(* IEC 61131-3 sources: volt/packages/volt-lsp-iec/test-corpus/bakon-nano/Device/Plc Logic/Application/Library Manager/Collections, 40 files *)

(* ---- PAIR_DINTDINT.dut ---- *)
TYPE PAIR_DINTDINT :
STRUCT
	DIKEY : DINT;
	DIVALUE : DINT;
END_STRUCT
END_TYPE

(* ---- PAIR_PSTRINGDINT.dut ---- *)
TYPE PAIR_PSTRINGDINT :
STRUCT
	PSTR : POINTER TO STRING;
	DI : DINT;
END_STRUCT
END_TYPE

(* ---- PAIR_PSTRINGXWORD.dut ---- *)
TYPE PAIR_PSTRINGXWORD :
STRUCT
	PSTR : POINTER TO STRING;
	XW : __XWORD;
END_STRUCT
END_TYPE

(* ---- PAIR_STRINGDINT.dut ---- *)
TYPE PAIR_STRINGDINT :
STRUCT
	STR : STRING;
	DI : DINT;
END_STRUCT
END_TYPE

(* ---- PAIR_STRINGSTRING.dut ---- *)
TYPE PAIR_STRINGSTRING :
STRUCT
	STRKEY : STRING;
	STRVALUE : STRING;
END_STRUCT
END_TYPE

(* ---- STATICMEMBUFFER.dut ---- *)
TYPE STATICMEMBUFFER :
STRUCT
	PDATA : POINTER TO BYTE;
	UDIDATASIZE : UDINT;
	XEXTENDDYNAMICALLY : BOOL;
END_STRUCT
END_TYPE

(* ---- GLOBALS.gvl ---- *)
VAR_GLOBAL
	COMPONENT_NAME : STRING := 'Collections';
	VECTOR_STRING_LEN : INT := 80;
	ERR_MB_ALREADY_ALLOCATED : UDINT := 16#2100;
	ERR_OK : UDINT := 0;
	ERR_PARAMETER : UDINT := 2;
	ERR_NOTINITIALIZED : UDINT := 3;
	ERR_NOBUFFER : UDINT := 6;
	ERR_NOTIMPLEMENTED : UDINT := 12;
	ERR_NO_OBJECT : UDINT := 16#16;
END_VAR

(* ---- GVL_DEBUGONLYCOLLECTIONS.gvl ---- *)
VAR_GLOBAL
	G_ST : STRING(255);
	G_PST : POINTER TO STRING(255);
END_VAR

(* ---- PSTRCAT.pou ---- *)
FUNCTION PSTRCAT : DINT
VAR_INPUT
	PSTDEST : POINTER TO STRING;
	PSTSRC : POINTER TO STRING;
	DIDESTSIZE : DINT;
END_VAR
END_FUNCTION

(* ---- PSTRCMP.pou ---- *)
FUNCTION PSTRCMP : INT
VAR_INPUT
	PSTR1 : POINTER TO STRING;
	PSTR2 : POINTER TO STRING;
END_VAR
END_FUNCTION

(* ---- PSTRICMP.pou ---- *)
FUNCTION PSTRICMP : INT
VAR_INPUT
	PSTR1 : POINTER TO STRING;
	PSTR2 : POINTER TO STRING;
END_VAR
END_FUNCTION

(* ---- PSTRIFIND.pou ---- *)
FUNCTION PSTRIFIND : INT
VAR_INPUT
	PST1 : POINTER TO STRING(255);
	PST2 : POINTER TO STRING(255);
END_VAR
END_FUNCTION

(* ---- PSTRLEN.pou ---- *)
FUNCTION PSTRLEN : DINT
VAR_INPUT
	PSTRING : POINTER TO STRING;
END_VAR
END_FUNCTION

(* ---- PSTRLENUNTIL.pou ---- *)
FUNCTION PSTRLENUNTIL : DINT
VAR_INPUT
	PST : POINTER TO STRING;
	STTOKENDELIMITERS : STRING;
END_VAR
END_FUNCTION

(* ---- PSTRTOUPPER.pou ---- *)
FUNCTION PSTRTOUPPER : STRING(255)
VAR_INPUT
	PSTVALUE : POINTER TO STRING(255);
END_VAR
END_FUNCTION

(* ---- ABSTRTREENODE.pou ---- *)
FUNCTION_BLOCK ABSTRTREENODE
VAR
	_FATHER : IBaseTreeNode;
	_ICOUNT : DINT;
	_IBASETREENODE : IBaseTreeNode;
	ABSTRNODETYPE : INT;
	CHILDCOUNT : DINT;
	PROCHILDREN : POINTER TO ARRAY [0..100] OF IBaseTreeNode;
	SORTED : BOOL;
END_VAR
END_FUNCTION_BLOCK

METHOD GETCHILD : IBaseTreeNode
VAR_INPUT
	DIINDEX : DINT;
END_VAR
END_METHOD

METHOD GETFATHER : IBaseTreeNode
END_METHOD

METHOD ABSTRCOMPARETO : INT
VAR_INPUT
	PSEARCHDATA : POINTER TO BYTE;
END_VAR
END_METHOD

METHOD PROFINDCHILDINDEX : DINT
VAR_INPUT
	PSEARCHDATA : POINTER TO BYTE;
END_VAR
END_METHOD

METHOD PROGETNODE : IBaseTreeNode
VAR_INPUT
	DIINDEX : DINT;
END_VAR
END_METHOD

METHOD PRVFINDBINARY : DINT
VAR_INPUT
	PSEARCHDATA : POINTER TO BYTE;
END_VAR
END_METHOD

METHOD PRVFINDLINEAR : DINT
VAR_INPUT
	PSEARCHDATA : POINTER TO BYTE;
END_VAR
END_METHOD

METHOD ADDREF : DINT
END_METHOD

METHOD FB_EXIT : BOOL
VAR_INPUT
	BINCOPYCODE : BOOL;
END_VAR
END_METHOD

METHOD FB_INIT : BOOL
VAR_INPUT
	BINITRETAINS : BOOL;
	BINCOPYCODE : BOOL;
END_VAR
END_METHOD

METHOD FB_REINIT : BOOL
END_METHOD

METHOD QUERYINTERFACE : POINTER TO POINTER TO BYTE
VAR_INPUT
	IID : DWORD;
	PRESULT : POINTER TO UDINT;
END_VAR
END_METHOD

METHOD RELEASE : DINT
END_METHOD

(* ---- BASEMAP.pou ---- *)
FUNCTION_BLOCK BASEMAP EXTENDS BaseVector
VAR
	_IUPDATECOUNT : INT;
	_BOPTIMIZEDSORTFORINSERTIONONLYATEND : BOOL;
	PROUSEOPTIMIZEDSORTFORINSERTIONATTHEEND : BOOL;
END_VAR
END_FUNCTION_BLOCK

METHOD BEGINUPDATE : UDINT
END_METHOD

METHOD ENDUPDATE : UDINT
END_METHOD

METHOD ABSTRCOMPARE : INT
VAR_INPUT
	PKEY1 : POINTER TO BYTE;
	PKEY2 : POINTER TO BYTE;
END_VAR
END_METHOD

METHOD ABSTRKEYPTRFROMINDEX : POINTER TO BYTE
VAR_INPUT
	UDIINDEX : UDINT;
END_VAR
END_METHOD

METHOD ABSTRSWAP : UDINT
VAR_INPUT
	INDEX1 : UDINT;
	INDEX2 : UDINT;
END_VAR
END_METHOD

METHOD PROADDMAPITEM : UDINT
VAR_INPUT
	PITEM : POINTER TO BYTE;
END_VAR
END_METHOD

METHOD PROFINDPAIRINDEX : DINT
VAR_INPUT
	PKEY : POINTER TO BYTE;
END_VAR
END_METHOD

METHOD PRVAFTERUPDATE : UDINT
VAR_INPUT
	BONLYSINGLEINSERT : BOOL;
END_VAR
END_METHOD

METHOD PRVBUBBLESORT : UDINT
END_METHOD

METHOD PRVCOMPAREBYINDEXANDVALUE : INT
VAR_INPUT
	UDI1 : UDINT;
	PKEYVAL : POINTER TO BYTE;
END_VAR
END_METHOD

METHOD PRVCOMPAREBYINDICES : INT
VAR_INPUT
	UDI1 : UDINT;
	UDI2 : UDINT;
END_VAR
END_METHOD

METHOD PRVINSERTIONSORTFORLAST : UDINT
END_METHOD

METHOD PRVSORT : UDINT
VAR_INPUT
	BONLYSINGLEINSERT : BOOL;
END_VAR
END_METHOD

(* ---- BASEVECTOR.pou ---- *)
FUNCTION_BLOCK BASEVECTOR
VAR
	_MEMORY : MemBuffer;
	_PDATA : POINTER TO ARRAY [0..100] OF DWORD;
	_DICURRENTALLOCSIZE : DINT;
	_DICURRENTINSERTPOSITION : DINT;
	CAPACITY : DINT;
	COUNT : DINT;
	PRODATAPTR : POINTER TO BYTE;
END_VAR
END_FUNCTION_BLOCK

METHOD CLEAR : UDINT
END_METHOD

METHOD INITMEMORY : UDINT
VAR_INPUT
	BUFFER : StaticMemBuffer;
END_VAR
END_METHOD

METHOD REMOVELAST : UDINT
END_METHOD

METHOD RESERVESPACE : UDINT
VAR_INPUT
	IITEMCOUNT : UDINT;
END_VAR
END_METHOD

METHOD ABSTRASSIGN : UDINT
VAR_INPUT
	PBT : POINTER TO BYTE;
	UDIINDEX : UDINT;
END_VAR
END_METHOD

METHOD ABSTRDATAPTRCHANGED : UDINT
END_METHOD

METHOD ABSTRGETELEMENTPTR : UDINT
VAR_INPUT
	UDIINDEX : UDINT;
END_VAR
VAR_OUTPUT
	PENTRY : POINTER TO BYTE;
END_VAR
END_METHOD

METHOD ABSTRSIZEOFELEMENT : UDINT
END_METHOD

METHOD PROADDITEM : UDINT
VAR_INPUT
	PBT : POINTER TO BYTE;
END_VAR
END_METHOD

METHOD PROAFTERALLOC
VAR_INPUT
	DIPREVALLOCSIZE : DINT;
	DICURRALLOCSIZE : DINT;
END_VAR
END_METHOD

METHOD PROREMOVE : UDINT
VAR_INPUT
	UDIINDEX : UDINT;
END_VAR
END_METHOD

METHOD PRVALLOC : UDINT
VAR_INPUT
	UDIITEMCOUNT : UDINT;
END_VAR
END_METHOD

(* ---- BRANCHNAMEDTREENODE.pou ---- *)
FUNCTION_BLOCK BRANCHNAMEDTREENODE EXTENDS NamedTreeNode
VAR
	_PCHILDREN : POINTER TO ARRAY [0..100] OF IBaseTreeNode;
	_ICHILDCOUNT : DINT;
	CHILDCOUNT : DINT;
	PROCHILDREN : POINTER TO ARRAY [0..100] OF IBaseTreeNode;
END_VAR
END_FUNCTION_BLOCK

(* ---- CASESENSITIVENAMEDTREENODE.pou ---- *)
FUNCTION_BLOCK CASESENSITIVENAMEDTREENODE EXTENDS NamedTreeNode
VAR
	CASESENSITIVECOMPARISON : BOOL;
END_VAR
END_FUNCTION_BLOCK

(* ---- DINTTODINTMAP.pou ---- *)
FUNCTION_BLOCK DINTTODINTMAP EXTENDS BaseMap
VAR
	_PITEMS : POINTER TO ARRAY [0..100] OF Pair_DintDint;
END_VAR
END_FUNCTION_BLOCK

METHOD ADDDINTPAIR : UDINT
VAR_INPUT
	DIKEY : DINT;
	DIVALUE : DINT;
END_VAR
END_METHOD

METHOD GETVALUE : DINT
VAR_INPUT
	DIKEY : DINT;
END_VAR
VAR_OUTPUT
	UDIRESULT : UDINT;
END_VAR
END_METHOD

METHOD ABSTRASSIGN : UDINT
VAR_INPUT
	PBT : POINTER TO BYTE;
	UDIINDEX : UDINT;
END_VAR
END_METHOD

METHOD ABSTRCOMPARE : INT
VAR_INPUT
	PKEY1 : POINTER TO BYTE;
	PKEY2 : POINTER TO BYTE;
END_VAR
END_METHOD

METHOD ABSTRDATAPTRCHANGED : UDINT
END_METHOD

METHOD ABSTRKEYPTRFROMINDEX : POINTER TO BYTE
VAR_INPUT
	UDIINDEX : UDINT;
END_VAR
END_METHOD

METHOD ABSTRSIZEOFELEMENT : UDINT
END_METHOD

METHOD ABSTRSWAP : UDINT
VAR_INPUT
	INDEX1 : UDINT;
	INDEX2 : UDINT;
END_VAR
END_METHOD

(* ---- DINTVECTOR.pou ---- *)
FUNCTION_BLOCK DINTVECTOR EXTENDS BaseVector
VAR
	_PARRDINT : POINTER TO ARRAY [0..100] OF DINT;
END_VAR
END_FUNCTION_BLOCK

METHOD ADDDINT : UDINT
VAR_INPUT
	ITEM : DINT;
END_VAR
END_METHOD

METHOD GETDINT : DWORD
VAR_INPUT
	UDIINDEX : UDINT;
END_VAR
VAR_OUTPUT
	UDIRESULT : UDINT;
END_VAR
END_METHOD

METHOD ABSTRASSIGN : UDINT
VAR_INPUT
	PBT : POINTER TO BYTE;
	UDIINDEX : UDINT;
END_VAR
END_METHOD

METHOD ABSTRDATAPTRCHANGED : UDINT
END_METHOD

METHOD ABSTRSIZEOFELEMENT : UDINT
END_METHOD

(* ---- DWORDVECTOR.pou ---- *)
FUNCTION_BLOCK DWORDVECTOR EXTENDS BaseVector
VAR
	_PARRDW : POINTER TO ARRAY [0..100] OF DWORD;
END_VAR
END_FUNCTION_BLOCK

METHOD ADDDWORD : UDINT
VAR_INPUT
	ITEM : DWORD;
END_VAR
END_METHOD

METHOD GETDWORD : DWORD
VAR_INPUT
	UDIINDEX : UDINT;
END_VAR
VAR_OUTPUT
	UDIRESULT : UDINT;
END_VAR
END_METHOD

METHOD REMOVE : UDINT
VAR_INPUT
	UDIINDEX : UDINT;
END_VAR
END_METHOD

METHOD ABSTRASSIGN : UDINT
VAR_INPUT
	PBT : POINTER TO BYTE;
	UDIINDEX : UDINT;
END_VAR
END_METHOD

METHOD ABSTRDATAPTRCHANGED : UDINT
END_METHOD

METHOD ABSTRGETELEMENTPTR : UDINT
VAR_INPUT
	UDIINDEX : UDINT;
END_VAR
VAR_OUTPUT
	PENTRY : POINTER TO BYTE;
END_VAR
END_METHOD

METHOD ABSTRSIZEOFELEMENT : UDINT
END_METHOD

(* ---- INSTANCEPATHBUILDINGBRANCHNODE.pou ---- *)
FUNCTION_BLOCK INSTANCEPATHBUILDINGBRANCHNODE EXTENDS InstancePathBuildingNode
VAR
	_PCHILDREN : POINTER TO ARRAY [0..100] OF IBaseTreeNode;
	_ICHILDCOUNT : DINT;
	_TYPE : InstancePathBuildingNodeType;
	CHILDCOUNT : DINT;
	INSTANCEPATHNODETYPE : InstancePathBuildingNodeType;
	PROCHILDREN : POINTER TO ARRAY [0..100] OF IBaseTreeNode;
END_VAR
END_FUNCTION_BLOCK

(* ---- INSTANCEPATHBUILDINGNODE.pou ---- *)
FUNCTION_BLOCK INSTANCEPATHBUILDINGNODE EXTENDS NamedTreeNode
VAR
	_IINSTANCEPATHBUILDINGNODE : IInstancePathBuildingNode;
	INSTANCEPATHNODETYPE : InstancePathBuildingNodeType;
	PRVFATHERASINSTANCEBUILDINGNODE : IInstancePathBuildingNode;
END_VAR
END_FUNCTION_BLOCK

METHOD GETFULLPATH : DINT
VAR_INPUT
	PBUFFER : POINTER TO STRING;
	DIBUFFERSIZE : DINT;
END_VAR
END_METHOD

METHOD PRVDOGETFULLPATH : DINT
VAR_INPUT
	PBUFFER : POINTER TO STRING;
	DIBUFFERSIZE : DINT;
END_VAR
END_METHOD

METHOD QUERYINTERFACE : POINTER TO POINTER TO BYTE
VAR_INPUT
	IID : DWORD;
	PRESULT : POINTER TO UDINT;
END_VAR
END_METHOD

(* ---- INSTANCEPATHNODEFINDER.pou ---- *)
FUNCTION_BLOCK INSTANCEPATHNODEFINDER
VAR
	_ROOTNODES : POINTER TO ARRAY [0..0] OF IBaseTreeNode;
	_ROOTNODECOUNT : DINT;
	PROROOTNODECOUNT : DINT;
	PROROOTNODES : POINTER TO ARRAY [0..100] OF IBaseTreeNode;
	PROTCALLNODEFOUNDFORROOTNODE : BOOL;
	PROTCALLNODENOTFOUNDFORROOTNODE : BOOL;
END_VAR
END_FUNCTION_BLOCK

METHOD FIND : IInstancePathBuildingNode
VAR_INPUT
	STPATH : STRING(255);
END_VAR
END_METHOD

METHOD FINDLONG : IInstancePathBuildingNode
VAR_INPUT
	PSTPATH : POINTER TO STRING;
END_VAR
END_METHOD

METHOD FINDLONGWITHDATA : IInstancePathBuildingNode
VAR_INPUT
	PSTPATH : POINTER TO STRING;
	PDATA : POINTER TO BYTE;
END_VAR
VAR_OUTPUT
	BEND : BOOL;
	PRT : POINTER TO IInstancePathBuildingNode;
END_VAR
END_METHOD

METHOD FINDWITHDATA : IInstancePathBuildingNode
VAR_INPUT
	STPATH : STRING(255);
	PDATA : POINTER TO BYTE;
END_VAR
VAR_OUTPUT
	BEND : BOOL;
	PRT : POINTER TO InstancePathBuildingNode;
END_VAR
END_METHOD

METHOD INITIALIZE : BOOL
VAR_INPUT
	PROOTNODES : POINTER TO ARRAY [0..100] OF IBaseTreeNode;
	INODECOUNT : DINT;
END_VAR
END_METHOD

METHOD ABSTRIGNOREROOTNODE : BOOL
VAR_INPUT
	PNODE : IInstancePathBuildingNode;
	PDATA : POINTER TO BYTE;
END_VAR
END_METHOD

METHOD ABSTRNODEFOUND : IInstancePathBuildingNode
VAR_INPUT
	PNODE : IInstancePathBuildingNode;
	PDATA : POINTER TO BYTE;
	BDIRECTCHILDFOUND : BOOL;
END_VAR
END_METHOD

METHOD ABSTRNODENOTFOUND : IInstancePathBuildingNode
VAR_INPUT
	PPARENT : IInstancePathBuildingNode;
	PDATA : POINTER TO BYTE;
	PSTPATH : POINTER TO STRING;
END_VAR
VAR_IN_OUT
	IOFFSETINPATH : DINT;
END_VAR
END_METHOD

METHOD ABSTRNOTFOUND : IInstancePathBuildingNode
VAR_INPUT
	PSTPATH : POINTER TO STRING;
END_VAR
END_METHOD

(* ---- MEMBUFFER.pou ---- *)
FUNCTION_BLOCK MEMBUFFER
VAR
	_MEMBUF : StaticMemBuffer;
	_BDYNAMIC : BOOL;
	_UDIALLOCATEDSIZE : UDINT;
	_PALLOCATEDDATA : POINTER TO BYTE;
END_VAR
END_FUNCTION_BLOCK

METHOD ALLOC : POINTER TO BYTE
VAR_INPUT
	UDISIZE : UDINT;
END_VAR
VAR_OUTPUT
	UDIRESULT : UDINT;
END_VAR
END_METHOD

METHOD CANRESIZE : BOOL
VAR_INPUT
	UDINEWSIZE : UDINT;
END_VAR
END_METHOD

METHOD FB_EXIT : UDINT
VAR_INPUT
	BINCOPYCODE : BOOL;
END_VAR
END_METHOD

METHOD INITSTATIC : UDINT
VAR_INPUT
	BUFFER : StaticMemBuffer;
END_VAR
END_METHOD

METHOD RESIZE : POINTER TO BYTE
VAR_INPUT
	UDINEWSIZE : UDINT;
END_VAR
VAR_OUTPUT
	UDIRESULT : UDINT;
END_VAR
END_METHOD

(* ---- NAMEDTREENODE.pou ---- *)
FUNCTION_BLOCK NAMEDTREENODE EXTENDS AbstrTreeNode
VAR
	_PSTNAME : POINTER TO STRING;
	_INAMEDTREENODE : INamedTreeNode;
	CASESENSITIVECOMPARISON : BOOL;
	NAME : POINTER TO STRING;
END_VAR
END_FUNCTION_BLOCK

METHOD FB_INIT : BOOL
VAR_INPUT
	BINITRETAINS : BOOL;
	BINCOPYCODE : BOOL;
END_VAR
END_METHOD

METHOD FINDCHILDBYNAME : INamedTreeNode
VAR_INPUT
	STNAME : STRING(256);
END_VAR
END_METHOD

METHOD ABSTRCOMPARETO : INT
VAR_INPUT
	PSEARCHDATA : POINTER TO BYTE;
END_VAR
END_METHOD

METHOD QUERYINTERFACE : POINTER TO POINTER TO BYTE
VAR_INPUT
	IID : DWORD;
	PRESULT : POINTER TO UDINT;
END_VAR
END_METHOD

(* ---- PSTRINGTODINTMAP.pou ---- *)
FUNCTION_BLOCK PSTRINGTODINTMAP EXTENDS BaseMap
VAR
	_PITEMS : POINTER TO ARRAY [0..100] OF Pair_PStringDint;
	_BCASESENSITIVE : BOOL := TRUE;
	_BCOPYSTRINGS : BOOL := FALSE;
	CASESENSITIVE : BOOL;
	COPYSTRINGS : BOOL;
END_VAR
END_FUNCTION_BLOCK

METHOD ADDPSTRINGDINTPAIR : UDINT
VAR_INPUT
	PSTR : POINTER TO STRING;
	DIVALUE : DINT;
END_VAR
END_METHOD

METHOD CLEAR : UDINT
END_METHOD

METHOD FB_EXIT : UDINT
VAR_INPUT
	BINCOPYCODE : BOOL;
END_VAR
END_METHOD

METHOD GETINDEX : DINT
VAR_INPUT
	PSTR : POINTER TO STRING;
END_VAR
VAR_OUTPUT
	UDIRESULT : UDINT;
END_VAR
END_METHOD

METHOD GETKEYBYINDEX : POINTER TO BYTE
VAR_INPUT
	UDIINDEX : UDINT;
END_VAR
VAR_OUTPUT
	UDIRESULT : UDINT;
END_VAR
END_METHOD

METHOD GETVALUE : DINT
VAR_INPUT
	PSTR : POINTER TO STRING;
END_VAR
VAR_OUTPUT
	UDIRESULT : UDINT;
END_VAR
END_METHOD

METHOD GETVALUEBYINDEX : DINT
VAR_INPUT
	UDIINDEX : UDINT;
END_VAR
VAR_OUTPUT
	UDIRESULT : UDINT;
END_VAR
END_METHOD

METHOD REMOVE : UDINT
VAR_INPUT
	UDIINDEX : UDINT;
END_VAR
END_METHOD

METHOD SETVALUEBYINDEX : UDINT
VAR_INPUT
	UDIINDEX : UDINT;
	DIVALUE : DINT;
END_VAR
END_METHOD

METHOD ABSTRASSIGN : UDINT
VAR_INPUT
	PBT : POINTER TO BYTE;
	UDIINDEX : UDINT;
END_VAR
END_METHOD

METHOD ABSTRCOMPARE : INT
VAR_INPUT
	PKEY1 : POINTER TO BYTE;
	PKEY2 : POINTER TO BYTE;
END_VAR
END_METHOD

METHOD ABSTRDATAPTRCHANGED : UDINT
END_METHOD

METHOD ABSTRGETELEMENTPTR : UDINT
VAR_INPUT
	UDIINDEX : UDINT;
END_VAR
VAR_OUTPUT
	PENTRY : POINTER TO BYTE;
END_VAR
END_METHOD

METHOD ABSTRKEYPTRFROMINDEX : POINTER TO BYTE
VAR_INPUT
	UDIINDEX : UDINT;
END_VAR
END_METHOD

METHOD ABSTRSIZEOFELEMENT : UDINT
END_METHOD

METHOD ABSTRSWAP : UDINT
VAR_INPUT
	INDEX1 : UDINT;
	INDEX2 : UDINT;
END_VAR
END_METHOD

(* ---- PSTRINGTOXWORDMAP.pou ---- *)
FUNCTION_BLOCK PSTRINGTOXWORDMAP EXTENDS BaseMap
VAR
	_PITEMS : POINTER TO ARRAY [0..100] OF Pair_PStringXWORD;
	_BCASESENSITIVE : BOOL := TRUE;
	_BCOPYSTRINGS : BOOL := FALSE;
	CASESENSITIVE : BOOL;
	COPYSTRINGS : BOOL;
END_VAR
END_FUNCTION_BLOCK

METHOD ADDPSTRINGXWORDPAIR : UDINT
VAR_INPUT
	PSTR : POINTER TO STRING;
	XW : __XWORD;
END_VAR
END_METHOD

METHOD CLEAR : UDINT
END_METHOD

METHOD FB_EXIT : UDINT
VAR_INPUT
	BINCOPYCODE : BOOL;
END_VAR
END_METHOD

METHOD GETINDEX : DINT
VAR_INPUT
	PSTR : POINTER TO STRING;
END_VAR
VAR_OUTPUT
	UDIRESULT : UDINT;
END_VAR
END_METHOD

METHOD GETKEYBYINDEX : POINTER TO BYTE
VAR_INPUT
	UDIINDEX : UDINT;
END_VAR
VAR_OUTPUT
	UDIRESULT : UDINT;
END_VAR
END_METHOD

METHOD GETVALUE : __XWORD
VAR_INPUT
	PSTR : POINTER TO STRING;
END_VAR
VAR_OUTPUT
	UDIRESULT : UDINT;
END_VAR
END_METHOD

METHOD GETVALUEBYINDEX : __XWORD
VAR_INPUT
	UDIINDEX : UDINT;
END_VAR
VAR_OUTPUT
	UDIRESULT : UDINT;
END_VAR
END_METHOD

METHOD REMOVE : UDINT
VAR_INPUT
	UDIINDEX : UDINT;
END_VAR
END_METHOD

METHOD SETVALUEBYINDEX : UDINT
VAR_INPUT
	UDIINDEX : UDINT;
	XW : __XWORD;
END_VAR
END_METHOD

METHOD ABSTRASSIGN : UDINT
VAR_INPUT
	PBT : POINTER TO BYTE;
	UDIINDEX : UDINT;
END_VAR
END_METHOD

METHOD ABSTRCOMPARE : INT
VAR_INPUT
	PKEY1 : POINTER TO BYTE;
	PKEY2 : POINTER TO BYTE;
END_VAR
END_METHOD

METHOD ABSTRDATAPTRCHANGED : UDINT
END_METHOD

METHOD ABSTRGETELEMENTPTR : UDINT
VAR_INPUT
	UDIINDEX : UDINT;
END_VAR
VAR_OUTPUT
	PENTRY : POINTER TO BYTE;
END_VAR
END_METHOD

METHOD ABSTRKEYPTRFROMINDEX : POINTER TO BYTE
VAR_INPUT
	UDIINDEX : UDINT;
END_VAR
END_METHOD

METHOD ABSTRSIZEOFELEMENT : UDINT
END_METHOD

METHOD ABSTRSWAP : UDINT
VAR_INPUT
	INDEX1 : UDINT;
	INDEX2 : UDINT;
END_VAR
END_METHOD

(* ---- PSTRINGVECTOR.pou ---- *)
FUNCTION_BLOCK PSTRINGVECTOR EXTENDS BaseVector
VAR
	_PARRPSTRINGS : POINTER TO ARRAY [0..100] OF POINTER TO STRING;
END_VAR
END_FUNCTION_BLOCK

METHOD ADDSTRING : UDINT
VAR_INPUT
	PSTRING : POINTER TO STRING;
END_VAR
END_METHOD

METHOD GETSTRING : POINTER TO STRING
VAR_INPUT
	UDIINDEX : UDINT;
END_VAR
VAR_OUTPUT
	UDIRESULT : UDINT;
END_VAR
END_METHOD

METHOD ABSTRASSIGN : UDINT
VAR_INPUT
	PBT : POINTER TO BYTE;
	UDIINDEX : UDINT;
END_VAR
END_METHOD

METHOD ABSTRDATAPTRCHANGED : UDINT
END_METHOD

METHOD ABSTRSIZEOFELEMENT : UDINT
END_METHOD

(* ---- SORTEDBRANCHNAMEDTREENODE.pou ---- *)
FUNCTION_BLOCK SORTEDBRANCHNAMEDTREENODE EXTENDS BranchNamedTreeNode
VAR
	SORTED : BOOL;
END_VAR
END_FUNCTION_BLOCK

(* ---- SORTEDINSTANCEPATHBUILDINGBRANCHNODE.pou ---- *)
FUNCTION_BLOCK SORTEDINSTANCEPATHBUILDINGBRANCHNODE EXTENDS InstancePathBuildingBranchNode
VAR
	SORTED : BOOL;
END_VAR
END_FUNCTION_BLOCK

(* ---- SORTEDPSTRINGVECTOR.pou ---- *)
FUNCTION_BLOCK SORTEDPSTRINGVECTOR EXTENDS BaseMap
VAR
	_PPITEMS : POINTER TO POINTER TO BYTE;
	_BCASESENSITIVE : BOOL;
	CASESENSITIVE : BOOL;
END_VAR
END_FUNCTION_BLOCK

METHOD ADDPSTRING : UDINT
VAR_INPUT
	PSTTEXT : POINTER TO BYTE;
END_VAR
END_METHOD

METHOD GETPSTRING : POINTER TO BYTE
VAR_INPUT
	DIINDEX : DINT;
END_VAR
VAR_OUTPUT
	UDIRESULT : UDINT;
END_VAR
END_METHOD

METHOD ABSTRASSIGN : UDINT
VAR_INPUT
	PBT : POINTER TO BYTE;
	UDIINDEX : UDINT;
END_VAR
END_METHOD

METHOD ABSTRCOMPARE : INT
VAR_INPUT
	PKEY1 : POINTER TO BYTE;
	PKEY2 : POINTER TO BYTE;
END_VAR
END_METHOD

METHOD ABSTRDATAPTRCHANGED : UDINT
END_METHOD

METHOD ABSTRGETELEMENTPTR : UDINT
VAR_INPUT
	UDIINDEX : UDINT;
END_VAR
VAR_OUTPUT
	PENTRY : POINTER TO BYTE;
END_VAR
END_METHOD

METHOD ABSTRKEYPTRFROMINDEX : POINTER TO BYTE
VAR_INPUT
	UDIINDEX : UDINT;
END_VAR
END_METHOD

METHOD ABSTRSIZEOFELEMENT : UDINT
END_METHOD

METHOD ABSTRSWAP : UDINT
VAR_INPUT
	INDEX1 : UDINT;
	INDEX2 : UDINT;
END_VAR
END_METHOD

(* ---- STRINGBUILDER.pou ---- *)
FUNCTION_BLOCK STRINGBUILDER
VAR
	_MEMORY : MemBuffer;
	_UDICURRENTSIZE : UDINT;
	_UDICURRENTALLOCSIZE : UDINT;
	_PDATA : POINTER TO BYTE;
	CAPACITY : UDINT;
	LENGTH : UDINT;
END_VAR
END_FUNCTION_BLOCK

METHOD APPENDCHAR : UDINT
VAR_INPUT
	C : BYTE;
END_VAR
END_METHOD

METHOD APPENDPSTRING : UDINT
VAR_INPUT
	PST : POINTER TO BYTE;
END_VAR
END_METHOD

METHOD APPENDSTRING : UDINT
VAR_INPUT
	STR : STRING;
END_VAR
END_METHOD

METHOD CLEAR
END_METHOD

METHOD GETPSTRINGRESULT : POINTER TO BYTE
END_METHOD

METHOD INITMEMORY : UDINT
VAR_INPUT
	BUFFER : StaticMemBuffer;
END_VAR
END_METHOD

METHOD RESERVESPACE : UDINT
VAR_INPUT
	UDINEWSIZE : UDINT;
END_VAR
END_METHOD

METHOD PRVALLOC : UDINT
VAR_INPUT
	UDINEWSIZE : UDINT;
END_VAR
END_METHOD

METHOD PRVAPPEND : UDINT
VAR_INPUT
	PST : POINTER TO BYTE;
	ILEN : DINT;
END_VAR
END_METHOD

METHOD PRVASSUREADDITIONALSIZE : UDINT
VAR_INPUT
	UDIADDSIZE : UDINT;
END_VAR
END_METHOD

(* ---- STRINGTODINTMAP.pou ---- *)
FUNCTION_BLOCK STRINGTODINTMAP EXTENDS BaseMap
VAR
	_PITEMS : POINTER TO ARRAY [0..100] OF Pair_StringDint;
	_BCASESENSITIVE : BOOL := TRUE;
	CASESENSITIVE : BOOL;
END_VAR
END_FUNCTION_BLOCK

METHOD ADDSTRINGDINTPAIR : UDINT
VAR_INPUT
	STR : STRING;
	DIVALUE : DINT;
END_VAR
END_METHOD

METHOD GETVALUE : DINT
VAR_INPUT
	STR : STRING;
END_VAR
VAR_OUTPUT
	UDIRESULT : UDINT;
END_VAR
END_METHOD

METHOD ABSTRASSIGN : UDINT
VAR_INPUT
	PBT : POINTER TO BYTE;
	UDIINDEX : UDINT;
END_VAR
END_METHOD

METHOD ABSTRCOMPARE : INT
VAR_INPUT
	PKEY1 : POINTER TO BYTE;
	PKEY2 : POINTER TO BYTE;
END_VAR
END_METHOD

METHOD ABSTRDATAPTRCHANGED : UDINT
END_METHOD

METHOD ABSTRKEYPTRFROMINDEX : POINTER TO BYTE
VAR_INPUT
	UDIINDEX : UDINT;
END_VAR
END_METHOD

METHOD ABSTRSIZEOFELEMENT : UDINT
END_METHOD

METHOD ABSTRSWAP : UDINT
VAR_INPUT
	INDEX1 : UDINT;
	INDEX2 : UDINT;
END_VAR
END_METHOD

(* ---- STRINGTOSTRINGMAP.pou ---- *)
FUNCTION_BLOCK STRINGTOSTRINGMAP EXTENDS BaseMap
VAR
	_PITEMS : POINTER TO ARRAY [0..100] OF Pair_StringString;
	_BCASESENSITIVE : BOOL := TRUE;
	CASESENSITIVE : BOOL;
END_VAR
END_FUNCTION_BLOCK

METHOD ADDSTRINGSTRINGPAIR : UDINT
VAR_INPUT
	STRKEY : STRING;
	STRVALUE : STRING;
END_VAR
END_METHOD

METHOD GETVALUE : STRING
VAR_INPUT
	STR : STRING;
END_VAR
VAR_OUTPUT
	UDIRESULT : UDINT;
END_VAR
END_METHOD

METHOD ABSTRASSIGN : UDINT
VAR_INPUT
	PBT : POINTER TO BYTE;
	UDIINDEX : UDINT;
END_VAR
END_METHOD

METHOD ABSTRCOMPARE : INT
VAR_INPUT
	PKEY1 : POINTER TO BYTE;
	PKEY2 : POINTER TO BYTE;
END_VAR
END_METHOD

METHOD ABSTRDATAPTRCHANGED : UDINT
END_METHOD

METHOD ABSTRKEYPTRFROMINDEX : POINTER TO BYTE
VAR_INPUT
	UDIINDEX : UDINT;
END_VAR
END_METHOD

METHOD ABSTRSIZEOFELEMENT : UDINT
END_METHOD

METHOD ABSTRSWAP : UDINT
VAR_INPUT
	INDEX1 : UDINT;
	INDEX2 : UDINT;
END_VAR
END_METHOD

(* ---- STRINGVECTOR.pou ---- *)
FUNCTION_BLOCK STRINGVECTOR EXTENDS BaseVector
VAR
	_PARRSTRINGS : POINTER TO ARRAY [0..100] OF STRING(VECTOR_STRING_LEN);
END_VAR
END_FUNCTION_BLOCK

METHOD ADDSTRING : UDINT
VAR_INPUT
	STRVAL : STRING(VECTOR_STRING_LEN);
END_VAR
END_METHOD

METHOD GETSTRING : STRING(VECTOR_STRING_LEN)
VAR_INPUT
	UDIINDEX : UDINT;
END_VAR
VAR_OUTPUT
	UDIRESULT : UDINT;
END_VAR
END_METHOD

METHOD REMOVEAT : UDINT
VAR_INPUT
	UDIINDEX : UDINT;
END_VAR
END_METHOD

METHOD ABSTRASSIGN : UDINT
VAR_INPUT
	PBT : POINTER TO BYTE;
	UDIINDEX : UDINT;
END_VAR
END_METHOD

METHOD ABSTRDATAPTRCHANGED : UDINT
END_METHOD

METHOD ABSTRGETELEMENTPTR : UDINT
VAR_INPUT
	UDIINDEX : UDINT;
END_VAR
VAR_OUTPUT
	PENTRY : POINTER TO BYTE;
END_VAR
END_METHOD

METHOD ABSTRSIZEOFELEMENT : UDINT
END_METHOD

(* ---- UTILTOKENIZER.pou ---- *)
FUNCTION_BLOCK UTILTOKENIZER
VAR
	_PSTRTOTOKENIZE : POINTER TO STRING;
	_PSTRTOTOKENIZEASBYTES : POINTER TO BYTE;
	_STRDELIMS : STRING;
	_INUMDELIMS : INT;
	_ICURRENTPOS : INT;
	_ISTRTOTOKENIZELEN : DINT;
	CURRENTPOSITION : INT;
END_VAR
END_FUNCTION_BLOCK

METHOD INITIALIZE : BOOL
VAR_INPUT
	PSTR : POINTER TO STRING;
	STRDELIMS : STRING;
END_VAR
END_METHOD

METHOD NEXTTOKEN : STRING(256)
VAR_OUTPUT
	BEND : BOOL;
	ITOKENSTARTOFFSET : DINT;
	ITOKENENDOFFSET : DINT;
END_VAR
END_METHOD

(* ---- XWORDVECTOR.pou ---- *)
FUNCTION_BLOCK XWORDVECTOR EXTENDS BaseVector
VAR
	_PARRXW : POINTER TO ARRAY [0..100] OF __XWORD;
END_VAR
END_FUNCTION_BLOCK

METHOD ADDXWORD : UDINT
VAR_INPUT
	ITEM : __XWORD;
END_VAR
END_METHOD

METHOD FB_EXIT
VAR_INPUT
	BINCOPYCODE : BOOL;
END_VAR
END_METHOD

METHOD GETXWORD : __XWORD
VAR_INPUT
	UDIINDEX : UDINT;
END_VAR
VAR_OUTPUT
	UDIRESULT : UDINT;
END_VAR
END_METHOD

METHOD REMOVE : UDINT
VAR_INPUT
	UDIINDEX : UDINT;
END_VAR
END_METHOD

METHOD ABSTRASSIGN : UDINT
VAR_INPUT
	PBT : POINTER TO BYTE;
	UDIINDEX : UDINT;
END_VAR
END_METHOD

METHOD ABSTRDATAPTRCHANGED : UDINT
END_METHOD

METHOD ABSTRGETELEMENTPTR : UDINT
VAR_INPUT
	UDIINDEX : UDINT;
END_VAR
VAR_OUTPUT
	PENTRY : POINTER TO BYTE;
END_VAR
END_METHOD

METHOD ABSTRSIZEOFELEMENT : UDINT
END_METHOD
